Fanuc KAREL source: KT00457.KL

PROGRAM KT00457
%NOLOCKGROUP
VAR
  P1: POSITION
  P2: XYZWPREXT
  OUT: BOOLEAN
BEGIN
    P2.Y = 2.0
  OUT = P1 >= P2
END KT00457
